PROGRAM MAIN
VAR
    Cell : FB_CartonCell := (Name := 'Carton Cell');
END_VAR

Cell.RunScan();

END_PROGRAM

(* stored: Version 1.1.0.1, ProductVersion 3.1.4024.53
   POU MAIN: Id {52592E20-A431-4FDA-93CC-000000000027} *)
